(* IEC 61131-3 sources: plcassist-cli/packages/volt-lsp-iec/test-corpus/lenze-mid/Device/Plc Logic/Application/Library Manager/CAA CANopen Stack, 4 files *)

(* ---- OBJECTDICTIONARY.gvl ---- *)
VAR_GLOBAL
	GC_UISTATE_IDX : UINT := 16#1F82;
	GC_UICANOPEN_KERNEL_STATE_IDX : UINT := 16#2001;
	GC_USICANOPEN_KERNEL_STATE_SUBIDX : USINT := 1;
	GC_UIEMCY_DEV_IDX : UINT := 16#2002;
	GC_UIEMCY_IDX : UINT := 16#2003;
	GC_UIEMCY_SUBIDX : USINT := 1;
	GC_UIPERMITSDOTRANSMISSION_IDX : UINT := 16#2004;
	GC_UISDOCHANNELLIMIT_IDX : UINT := 16#2005;
	GC_UIBLOCKFDTACCESS_IDX : UINT := 16#2006;
END_VAR

(* ---- VERSIONCONSTANTS.gvl ---- *)
VAR_GLOBAL
	GC_BYVERSION : BYTE := 1;
	GC_BYVERSION_1 : BYTE := 0;
END_VAR

(* ---- ICANOPENSTACK.itf ---- *)
INTERFACE ICANOPENSTACK
END_INTERFACE

METHOD SDOABORT : PROC_STATE
VAR_INPUT
	ECMD : PROC_CMD;
	PPARAM : POINTER TO SDO_ABORT;
END_VAR
VAR_OUTPUT
	EERROR : ERROR;
END_VAR
END_METHOD

METHOD SDOWRITE : PROC_STATE
VAR_INPUT
	ECMD : PROC_CMD;
	PPARAM : POINTER TO SDO_WRITE;
END_VAR
VAR_OUTPUT
	EERROR : ERROR;
END_VAR
END_METHOD

METHOD SDOREAD : PROC_STATE
VAR_INPUT
	ECMD : PROC_CMD;
	PPARAM : POINTER TO SDO_READ;
END_VAR
VAR_OUTPUT
	EERROR : ERROR;
END_VAR
END_METHOD

METHOD STKOPEN : PROC_STATE
VAR_INPUT
	ECMD : PROC_CMD;
	USINETID : USINT;
	USINODEID : USINT;
	UIBAUDRATE : UINT;
	ESPEC : STK_SPEC;
END_VAR
VAR_OUTPUT
	EERROR : ERROR;
END_VAR
END_METHOD

METHOD STKCLOSE : PROC_STATE
VAR_INPUT
	ECMD : PROC_CMD;
END_VAR
VAR_OUTPUT
	EERROR : ERROR;
END_VAR
END_METHOD

METHOD STKGETINFO : PROC_STATE
VAR_INPUT
	ECMD : PROC_CMD;
	PSTKINFO : POINTER TO STK_INFO;
	PNETINFO : POINTER TO NET_INFO;
END_VAR
VAR_OUTPUT
	EERROR : ERROR;
END_VAR
END_METHOD

(* ---- GETSUPPLIERVERSION.fun ---- *)
FUNCTION GETSUPPLIERVERSION : WORD
VAR_INPUT
	XDUMMY : BOOL;
END_VAR
END_FUNCTION
